(* This testsuite tests the function block FB_AdjustAssertFailureMessageToMax255CharLength_Test
   The total printed message can not be more than 253 characters long.
*)
FUNCTION_BLOCK FB_AdjustAssertFailureMessageToMax253CharLengthTest EXTENDS TcUnit.FB_TestSuite

TestInstancePath253CharsExpectTooLongTestInstancePath();
TestInstancePath221CharsExpectShortenedTestInstancePath();
TestInstancePath255CharsExpectTooLongTestInstancePath();

METHOD TestInstancePath221CharsExpectShortenedTestInstancePath
VAR
    AdjustAssertFailureMessageToMax253CharLength : FB_AdjustAssertFailureMessageToMax253CharLength;

    // @Text-Fixture
    TestInstancePathNameWith221Chars : T_MaxString := 'PRG_TEST.LongInstanceNameLongInstanceNameLongInstanceNameLongInstanceNameLongInstanceNameLongInstanceNameLongInstanceNameLongInstanceNameLongInstanceNameLongInstanceName@LONGTESTNAMELONGTESTNAMELONGTESTNAMELONGTESTNAMELON';
    TooLongTestMessage60Chars : T_MaxString := 'Very long message that is 60 characters long which means tha';

    // @Test-Result-Expected
    // 221 + 32 = 253 (in other words, expected test message should be 32 characters long including '...TestMsg too long'
    TestMessageResultExpected : T_MaxString := 'Very long mes...TestMsg too long'; 

    // @Test-Result
    TestInstancePathResult : T_MaxString;
    TestMessageResult : T_MaxString;
END_VAR
TEST('TestInstancePath221CharsExpectShortenedTestInstancePath');

AdjustAssertFailureMessageToMax253CharLength(TestInstancePath := TestInstancePathNameWith221Chars,
                                             TestMessage := TooLongTestMessage60Chars,
                                             TestInstancePathProcessed => TestInstancePathResult,
                                             TestMessageProcessed => TestMessageResult);


AssertEquals_STRING(Expected := TestInstancePathNameWith221Chars, // Same test instance path should be expected as the one going in
                    Actual := TestInstancePathResult,
                    'Test instance path not correct');

AssertEquals_STRING(Expected := TestMessageResultExpected,
                    Actual := TestMessageResult,
                    'Test message not correct');

TEST_FINISHED();
END_METHOD

METHOD PRIVATE TestInstancePath253CharsExpectTooLongTestInstancePath
VAR
    AdjustAssertFailureMessageToMax253CharLength : FB_AdjustAssertFailureMessageToMax253CharLength;

    // @Text-Fixture
    TestInstancePathNameWith253Chars : T_MaxString := 'PRG_TEST.LongInstanceNameLongInstanceNameLongInstanceNameLongInstanceNameLongInstanceNameLongInstanceNameLongInstanceNameLongInstanceNameLongInstanceNameLongInstanceName@LONGTESTNAMELONGTESTNAMELONGTESTNAMELONGTESTNAMELONGTESTNAMELONGTESTNAMELONGTESTNAM';
    ShortTestMessage : T_MaxString := 'Very short message';

    // @Test-Result-Expected
    TestInstancePathNameWith253CharsExpectedResult : T_MaxString := 'PRG_TEST.LongInstanceNameLongInstanceNameLongInstanceNameLongInstanceNameLongInstanceNameLongInstanceNameLongInstanceNameLongInstanceNameLongInstanceNameLongInstanceName@LONGTESTNAMELONGTESTNAMELONGTESTNAMELONGTESTNAMELONGTESTNAMELON...TestName too long';
    ShortTestMessageExpectedResult : T_MaxString := '';

    // @Test-Result
    TestInstancePathNameWith253CharsResult : T_MaxString;
    ShortTestMessageResult : T_MaxString;
END_VAR
TEST('TestInstancePath253CharsExpectTooLongTestInstancePath');

AdjustAssertFailureMessageToMax253CharLength(TestInstancePath := TestInstancePathNameWith253Chars,
                                             TestMessage := ShortTestMessage,
                                             TestInstancePathProcessed => TestInstancePathNameWith253CharsResult,
                                             TestMessageProcessed => ShortTestMessageResult);

AssertEquals_STRING(Expected := TestInstancePathNameWith253CharsExpectedResult,
                    Actual := TestInstancePathNameWith253CharsResult,
                    'Test instance path not correct');

AssertEquals_STRING(Expected := ShortTestMessageExpectedResult,
                    Actual := ShortTestMessageResult,
                    'Test message not correct');

TEST_FINISHED();
END_METHOD

METHOD PRIVATE TestInstancePath255CharsExpectTooLongTestInstancePath
VAR
    AdjustAssertFailureMessageToMax253CharLength : FB_AdjustAssertFailureMessageToMax253CharLength;

    // @Text-Fixture
    TestInstancePathNameWith255Chars : T_MaxString := 'PRG_TEST.LongInstanceNameLongInstanceNameLongInstanceNameLongInstanceNameLongInstanceNameLongInstanceNameLongInstanceNameLongInstanceNameLongInstanceNameLongInstanceName@LONGTESTNAMELONGTESTNAMELONGTESTNAMELONGTESTNAMELONGTESTNAMELONGTESTNAMELONGTESTNAGAV';
    ShortTestMessage : T_MaxString := 'Very short message';

    // @Test-Result-Expected
    TestInstancePathNameWith253CharsExpectedResult : T_MaxString := 'PRG_TEST.LongInstanceNameLongInstanceNameLongInstanceNameLongInstanceNameLongInstanceNameLongInstanceNameLongInstanceNameLongInstanceNameLongInstanceNameLongInstanceName@LONGTESTNAMELONGTESTNAMELONGTESTNAMELONGTESTNAMELONGTESTNAMELON...TestName too long';
    ShortTestMessageExpectedResult : T_MaxString := '';

    // @Test-Result
    TestInstancePathNameWith253CharsResult : T_MaxString;
    ShortTestMessageResult : T_MaxString;
END_VAR
TEST('TestInstancePath255CharsExpectTooLongTestInstancePath');

AdjustAssertFailureMessageToMax253CharLength(TestInstancePath := TestInstancePathNameWith255Chars,
                                             TestMessage := ShortTestMessage,
                                             TestInstancePathProcessed => TestInstancePathNameWith253CharsResult,
                                             TestMessageProcessed => ShortTestMessageResult);

AssertEquals_STRING(Expected := TestInstancePathNameWith253CharsExpectedResult,
                    Actual := TestInstancePathNameWith253CharsResult,
                    'Test instance path not correct');

AssertEquals_STRING(Expected := ShortTestMessageExpectedResult,
                    Actual := ShortTestMessageResult,
                    'Test message not correct');

TEST_FINISHED();
END_METHOD

END_FUNCTION_BLOCK

(* stored: Version 1.1.0.1
   POU FB_AdjustAssertFailureMessageToMax253CharLengthTest: Id {305341a5-f462-4bcb-ba17-ae2773c50e69}, SpecialFunc None
   Method TestInstancePath221CharsExpectShortenedTestInstancePath: Id {dc008964-f701-440f-97f6-bba60a51fe93}
   Method TestInstancePath253CharsExpectTooLongTestInstancePath: Id {f67e3ff5-02f7-4268-9fa7-f06935f8269a}
   Method TestInstancePath255CharsExpectTooLongTestInstancePath: Id {fbb2640b-9b30-45ae-a207-49da858d57e9} *)
